PROGRAM ContextFactory

(*
	Allocates a span context holding copies of the given identity. The caller owns pDest.
	The identifiers are not validated; producers are responsible for what they build,
	and a context built from all-zero identifiers is simply not valid.
	pTraceState is borrowed and copied; 0 means no trace state.
*)
METHOD buildContext : BOOL
VAR_IN_OUT
	pDest: POINTER TO FB_SpanContext;
END_VAR
VAR_INPUT
	pTraceId: POINTER TO FB_TraceId;
	pSpanId: POINTER TO FB_SpanId;
	pTraceState: POINTER TO FB_TraceState;
	traceFlags: UDINT;
END_VAR
VAR_OUTPUT
	failureReason: E_ContextFactoryFailureReason;
END_VAR
VAR
	_pTraceState: POINTER TO FB_TraceState;
	_pNew: POINTER TO FB_SpanContext;
END_VAR
buildContext := FALSE;
failureReason := E_ContextFactoryFailureReason.NA;

IF pDest <> 0 THEN
	failureReason := E_ContextFactoryFailureReason.DESTINATION_ALREADY_ASSIGNED;
	RETURN;
END_IF

IF pTraceId = 0 THEN
	failureReason := E_ContextFactoryFailureReason.TRACE_ID_POINTER_NULL;
	RETURN;
END_IF

IF pSpanId = 0 THEN
	failureReason := E_ContextFactoryFailureReason.SPAN_ID_POINTER_NULL;
	RETURN;
END_IF

// clone all owned data before allocating the context itself
IF pTraceState <> 0 THEN
	IF NOT TraceStateFactory.clone(pDest:=_pTraceState, pSrc:=pTraceState) THEN
		failureReason := E_ContextFactoryFailureReason.MEMORY_ALLOCATION_FAILURE;
		RETURN;
	END_IF
END_IF

_pNew := __NEW(FB_SpanContext(
	pTraceId:=pTraceId,
	pSpanId:=pSpanId,
	pTraceState:=_pTraceState,
	traceFlags:=traceFlags
));
IF _pNew = 0 THEN
	failureReason := E_ContextFactoryFailureReason.MEMORY_ALLOCATION_FAILURE;
	IF _pTraceState <> 0 THEN _pTraceState^.delete(pSelf:=_pTraceState); END_IF
	RETURN;
END_IF
_pTraceState := 0;  // moved into FB_SpanContext
pDest := _pNew;
buildContext := failureReason = E_ContextFactoryFailureReason.NA;
END_METHOD

(*
	Allocates a snapshot of a span's identity. The caller owns pDest, which must be 0; the span
	is borrowed and unchanged. The span is the producer, and its identifiers come from the id
	generator, which only hands out valid ones, so they are not checked again here. A span that
	has not been built has no identifiers and is refused with TRACE_ID_POINTER_NULL.
	The context is always local: a span's own flags describe its parent's remoteness, so only
	the W3C trace flags are kept, and remoteness is marked as known and not remote.
*)
METHOD fromSpan : BOOL
VAR_IN_OUT
	pDest: POINTER TO FB_SpanContext;
END_VAR
VAR_INPUT
	pSpan: POINTER TO FB_Span;
END_VAR
VAR_OUTPUT
	failureReason: E_ContextFactoryFailureReason;
END_VAR
VAR
	_traceFlags: UDINT;
END_VAR
fromSpan := FALSE;
failureReason := E_ContextFactoryFailureReason.NA;

IF pSpan = 0 THEN
	failureReason := E_ContextFactoryFailureReason.SPAN_POINTER_NULL;
	RETURN;
END_IF

_traceFlags := (pSpan^.flags AND TO_UDINT(E_SpanFlags.SPAN_FLAGS_TRACE_FLAGS_MASK))
	OR TO_UDINT(E_SpanFlags.SPAN_FLAGS_CONTEXT_HAS_IS_REMOTE_MASK);

fromSpan := ContextFactory.buildContext(
	pDest:=pDest,
	pTraceId:=pSpan^.traceId,
	pSpanId:=pSpan^.spanId,
	pTraceState:=pSpan^.traceState,
	traceFlags:=_traceFlags,
	failureReason=>failureReason
);
END_METHOD

END_PROGRAM

(* stored: Version 1.1.0.1
   POU ContextFactory: Id {63c02e55-2619-431c-a44a-88f22902c2e9}, SpecialFunc None
   Method buildContext: Id {d94b6c45-a4ff-4e52-afe3-b7fcb8bb8c8f}
   Method fromSpan: Id {f7f7f5f2-0b21-4cce-8675-bb1ea9059427} *)
